TYPE (* Data type with four variables *)
  (* Standard: 61499-1; Description: Copyright (c) 2023 Johannes Kepler University Linz This program and the accompanying materials are made available under the terms of the Eclipse Public License 2.0 which is available at https://www.eclipse.org/legal/epl-2.0/ SPDX-License-Identifier: EPL-2.0 *)
  (* Version 1.0, 2023-03-08, Bianca Wiesmayr, Johannes Kepler University Linz, initial API and implementation and/or initial documentation *)
  structtype : STRUCT
    VAR1 : BOOL := true;
    VAR2 : INT := INT#-5;
    VAR3 : UINT := UINT#17;
    VAR4 : WORD := 16#AFFE;
  END_STRUCT;
END_TYPE
